(*
SPDX-FileCopyrightText: © 2026 Oleksandr Tiutyk <trofimich@gmail.com>
SPDX-License-Identifier: MIT
License: https://opensource.org/license/mit
*)

(*!
<summary>Defines the execution outcome of an individual test scenario.</summary>
<description>
Tracks whether a test has not yet run, is currently executing across cycles, passed all assertions, failed an
assertion or invariant, or was explicitly skipped.
</description>
*)

{attribute 'qualified_only'}
{attribute 'strict'}
{attribute 'to_string'}
TYPE TEST_OUTCOME :
(
	NOT_RUN := 0,
	RUNNING := 1,
	PASSED := 2,
	FAILED := 3,
	SKIPPED := 4
);
END_TYPE

(* stored: Version 1.1.0.1
   DUT TEST_OUTCOME: Id {d0a3c1bd-065a-4382-9ec0-e018efd469c3} *)
